// TIA Portal V20 export
VAR_GLOBAL   // PLC tag table "Laser_in_macsa"
   "-XT500_d_counter" AT %ID1583 : DWord;   // counter indicating the number of o.k. prints since entering into the printing mode
   "-XT500_s_counter" AT %ID1587 : DWord;   // counter indicating the number of prints since entering into the printing mode.
   "-XT500_messageport" AT %ID1591 : DWord;   // indicates the bit combination of the external message selection (when external message mode is activated)
   "-XT500_status_byte_0" AT %IB1595 : Byte;
   "-XT500_status_byte_1" AT %IB1596 : Byte;   // 0x00: default value. -- 0x01: request; the system is requesting information to
   "-XT500_status_byte_2" AT %IB1597 : Byte;   // option byte; (internal use), indicates the type of
   "-XT500_status_byte_3" AT %IB1598 : Byte;   // 0x00: default , system is in standard mode. 0x01: system is in external message selection mode 0x04: system is in a batch-job mode.
   "-XT500_t_counter" AT %ID1599 : DWord;   // 32-bit counter indicating the total number of prints of the laser system
   "-XT500_copies" AT %ID1603 : DWord;   // the actual number of print copies.
   "-XT500_alarm_information" AT %IW1609 : Word;   // 0X0000: no alarms -- 0x0C0E: wrong messageport (no file found for the external message selection) -- 0x0848: alarms active; some alarms are active (interlock, shutter,....) -- 0xFFFF: initialization of the firmware has failed due to some hardware failure.
   "-XT500_prinntime" AT %ID1611 : DWord;   // print time
   "-XT500_alarm-mask" AT %ID1616 : DWord;   // popis panel text end grafik list
   "-XT500_signalstate" AT %ID1619 : DWord;
   "-XT500_name_byte_0" AT %IB1623 : Byte;   // actual filename + extension of the message.
   "-XT500_name_byte_1" AT %IB1624 : Byte;   // actual filename + extension of the message.
   "-XT500_name_byte_2" AT %IB1625 : Byte;   // actual filename + extension of the message.
   "-XT500_name_byte_3" AT %IB1626 : Byte;   // actual filename + extension of the message.
   "-XT500_name_byte_4" AT %IB1627 : Byte;   // actual filename + extension of the message.
   "-XT500_name_byte_5" AT %IB1628 : Byte;   // actual filename + extension of the message.
   "-XT500_name_byte_6" AT %IB1629 : Byte;   // actual filename + extension of the message.
   "-XT500_name_byte_7" AT %IB1630 : Byte;   // actual filename + extension of the message.
   "-XT500_name_byte_8" AT %IB1631 : Byte;   // actual filename + extension of the message.
   "-XT500_name_byte_9" AT %IB1632 : Byte;   // actual filename + extension of the message.
   "-XT500_name_byte_10" AT %IB1633 : Byte;   // actual filename + extension of the message.
   "-XT500_name_byte_11" AT %IB1634 : Byte;   // actual filename + extension of the message.
   "-XT500_name_byte_12" AT %IB1635 : Byte;   // actual filename + extension of the message.
   "-XT500_name_byte_13" AT %IB1636 : Byte;   // actual filename + extension of the message.
   "-XT500_name_byte_14" AT %IB1637 : Byte;   // actual filename + extension of the message.
   "-XT500_name_byte_15" AT %IB1638 : Byte;   // actual filename + extension of the message.
   "-XT500_eventhandler_byte_0" AT %IB1639 : Byte;   // actual filename + extension of the eventhandler-file.
   "-XT500_eventhandler_byte_1" AT %IB1640 : Byte;   // actual filename + extension of the eventhandler-file.
   "-XT500_eventhandler_byte_2" AT %IB1641 : Byte;   // actual filename + extension of the eventhandler-file.
   "-XT500_eventhandler_byte_3" AT %IB1642 : Byte;   // actual filename + extension of the eventhandler-file.
   "-XT500_eventhandler_byte_4" AT %IB1643 : Byte;   // actual filename + extension of the eventhandler-file.
   "-XT500_eventhandler_byte_5" AT %IB1644 : Byte;   // actual filename + extension of the eventhandler-file.
   "-XT500_eventhandler_byte_6" AT %IB1645 : Byte;   // actual filename + extension of the eventhandler-file.
   "-XT500_eventhandler_byte_7" AT %IB1646 : Byte;   // actual filename + extension of the eventhandler-file.
   "-XT500_eventhandler_byte_8" AT %IB1647 : Byte;   // actual filename + extension of the eventhandler-file.
   "-XT500_eventhandler_byte_9" AT %IB1648 : Byte;   // actual filename + extension of the eventhandler-file.
   "-XT500_eventhandler_byte_10" AT %IB1649 : Byte;   // actual filename + extension of the eventhandler-file.
   "-XT500_eventhandler_byte_11" AT %IB1650 : Byte;   // actual filename + extension of the eventhandler-file.
   "-XT500_eventhandler_byte_12" AT %IB1651 : Byte;   // actual filename + extension of the eventhandler-file.
   "-XT500_eventhandler_byte_13" AT %IB1652 : Byte;   // actual filename + extension of the eventhandler-file.
   "-XT500_eventhandler_byte_14" AT %IB1653 : Byte;   // actual filename + extension of the eventhandler-file.
   "-XT500_eventhandler_byte_15" AT %IB1654 : Byte;   // actual filename + extension of the eventhandler-file.
   "-XT500_extended_alarm-mask" AT %ID1655 : DWord;   // See Status command. When the alarm-mask has the ‘extended alarmmask’ rozepsano text list
   "-XT500_not_used_0" AT %IB1659 : Byte;
   "-XT500_not_used_1" AT %IB1660 : Byte;
   "-XT500_scanfield_0" AT %IB1661 : Byte;
   "-XT500_scanfield_1" AT %IB1662 : Byte;
   "-XT500_data_recived_byte" AT %IB1663 : Byte;   // status
   "-XT500_data_recived_byte_0" AT %I1663.0 : Bool;   // data ready
   "-XT500_data_recived_byte_1" AT %I1663.1 : Bool;   // clear command error trigger
   "-XT500_data_recived_byte_2" AT %I1663.2 : Bool;
   "-XT500_data_recived_byte_3" AT %I1663.3 : Bool;
   "-XT500_data_recived_byte_4" AT %I1663.4 : Bool;
   "-XT500_data_recived_byte_5" AT %I1663.5 : Bool;
   "-XT500_data_recived_byte_6" AT %I1663.6 : Bool;
   "-XT500_data_recived_byte_7" AT %I1663.7 : Bool;
   "-XT500_command_error_info" AT %IW1664 : Word;   // command error info (0xFF == command
   "-XT500_status_byte_0_bool_0" AT %I1595.0 : Bool;   // when set, system is in printing mode (waiting for photocell/PLC)
   "-XT500_status_byte_0_bool_1" AT %I1595.1 : Bool;   // when set, system is actually printing a message
   "-XT500_status_byte_0_bool_2" AT %I1595.2 : Bool;   // when set, system is waiting for a 'alarm reset' signal (DSP cards only).
   "-XT500_status_byte_0_bool_3" AT %I1595.3 : Bool;   // when set, system is waiting for an input signal (DSP cards only)
   "-XT500_status_byte_0_bool_4" AT %I1595.4 : Bool;   // when set, system is waiting for an external motorized axis to reach a new position.
   "-XT500_status_byte_0_bool_5" AT %I1595.5 : Bool;   // when set, system is in ‘printsession’ mode.
   "-XT500_status_byte_0_bool_6" AT %I1595.6 : Bool;   // reserved
   "-XT500_status_byte_0_bool_7" AT %I1595.7 : Bool;   // reserved
   "-XT500_status_byte_1_bool_0" AT %I1596.0 : Bool;
   "-XT500_status_byte_1_bool_1" AT %I1596.1 : Bool;
   "-XT500_status_byte_1_bool_2" AT %I1596.2 : Bool;
   "-XT500_status_byte_1_bool_3" AT %I1596.3 : Bool;
   "-XT500_status_byte_1_bool_4" AT %I1596.4 : Bool;
   "-XT500_status_byte_1_bool_5" AT %I1596.5 : Bool;
   "-XT500_status_byte_1_bool_6" AT %I1596.6 : Bool;
   "-XT500_status_byte_1_bool_7" AT %I1596.7 : Bool;
   "-XT500_scanfield_1_bit_8" AT %I1662.0 : Bool;
   "-XT500_scanfield_1_bit_9" AT %I1662.1 : Bool;
   "-XT500_scanfield_1_bit_10" AT %I1662.2 : Bool;   // 0: static
   "-XT500_scanfield_1_bit_11" AT %I1662.3 : Bool;   // 1: dynamic
   "-XT500_scanfield_1_bit_12" AT %I1662.4 : Bool;   // 2: dynamic-distance
   "-XT500_scanfield_1_bit_13" AT %I1662.5 : Bool;   // 3: static-dynamic
   "-XT500_scanfield_1_bit_14" AT %I1662.6 : Bool;   // 4: stepper mode
   "-XT500_scanfield_1_bit_15" AT %I1662.7 : Bool;   // 5: XY stepper mode
   "-XT500_alarm-mask_interlock" AT %I1618.0 : Bool;   // interlock součást alarm-mask
   "-XT500_alarm-mask_shutter" AT %I1618.3 : Bool;   // shutter součást alarm-mask oim
   "-XT500_alarm-mask_laser_not_ready" AT %I1618.4 : Bool;   // laser nor ready součást alarm mask
   "-XT500_alarm-mask_laser_not_armed" AT %I1619.3 : Bool;   // laser nor armed součást alarm mask
   "-XT500_alarm_mas_warm_up_in_progres" AT %I1619.5 : Bool;   // warm_up_in_progres součást alarm mask
   "-XT500_alarm-mask_shutter_oim" AT %I1618.1 : Bool;
   "-XT500_copies_1" AT %IW1605 : Word;
   "-XT500_copies_2" AT %IW1607 : Word;
   "-XT500_Tag_1" AT %I1618.2 : Bool;
   "-XT500_alarm_information(1)" AT %IW1610 : Word;   // 0X0000: no alarms -- 0x0C0E: wrong messageport (no file found for the external message selection) -- 0x0848: alarms active; some alarms are active (interlock, shutter,....) -- 0xFFFF: initialization of the firmware has failed due to some hardware failure.
   "-XT500_alarm_information(2)" AT %IW1608 : Word;   // 0X0000: no alarms -- 0x0C0E: wrong messageport (no file found for the external message selection) -- 0x0848: alarms active; some alarms are active (interlock, shutter,....) -- 0xFFFF: initialization of the firmware has failed due to some hardware failure.
   "-XT500_alarm_information(3)" AT %IW1611 : Word;   // 0X0000: no alarms -- 0x0C0E: wrong messageport (no file found for the external message selection) -- 0x0848: alarms active; some alarms are active (interlock, shutter,....) -- 0xFFFF: initialization of the firmware has failed due to some hardware failure.
   "-XT500_alarm_information_bool_1" AT %I1610.0 : Bool;
   "-XT500_alarm_information_bool_2" AT %I1610.1 : Bool;
   "-XT500_alarm_information_bool_3" AT %I1610.2 : Bool;
   "-XT500_alarm_information_bool_4" AT %I1610.3 : Bool;   // neni_nahrato_1
   "-XT500_alarm_information_bool_5" AT %I1610.4 : Bool;
   "-XT500_alarm_information_bool_6" AT %I1610.5 : Bool;
   "-XT500_alarm_information_bool_7" AT %I1610.6 : Bool;   // neni_najrato_2
   "-XT500_alarm_information_bool_8" AT %I1610.7 : Bool;
END_VAR
